Staubli VAL3: resetAlarm.pgx

public program resetAlarm()
  local num l_n
begin
  for l_n=0 to size(_nAlarmCode)-1
    _nErrIndex[l_n]=-1
    _nAlarmCode[l_n]=0
    sAlarmMes[l_n]=""
  endFor
  _nAlarmIndex=0
end
